(*
SPDX-FileCopyrightText: © 2026 Oleksandr Tiutyk <trofimich@gmail.com>
SPDX-License-Identifier: MIT
License: https://opensource.org/license/mit
*)

(*!
<summary>Provides an embedded variable reset scope for child condition attachment.</summary>
*)
{attribute 'hide'}
INTERFACE IVariableResetScopeProvider EXTENDS TOF_Core.IObject

(*!
<summary>Borrows the variable reset scope embedded in this parent for condition attachment.</summary>
<description>Returns live storage for the lifetime of the parent. Used by the validated parent setter
in its owning task. The caller must not delete, copy or independently reconfigure the scope.</description>
*)
METHOD GetResetScope : IVariableResetScope
END_METHOD

END_INTERFACE

(* stored: Version 1.1.0.1
   Itf IVariableResetScopeProvider: Id {b6f055fb-1303-40b6-ae46-be3e1197609f}
   Method GetResetScope: Id {ccb26761-efc3-472a-affa-9a148448d3a5} *)
